% RSLogix 500 project PROGRAM 4.RSS, saved by version 8.30.00.16 %
PROJECT "UNTITLED"    % processor: Bul.1763 MicroLogix 1100 Series B %

PROGRAM FILES
  LAD 2 "MAIN"  8 rungs
  LAD 3 "IO"  7 rungs
  LAD 4 "CONTROLS"  7 rungs
  LAD 5 "CYCL_CTRL"  5 rungs
  LAD 6 "SERVO_CTRL"  4 rungs
  LAD 7 "VALVE_CTRL"  7 rungs
  LAD 8 "POS_CTRL"  6 rungs
  LAD 9 "TIMERS"  4 rungs

DATA FILES
  O0 OUTPUT  4 elements
  I1 INPUT  6 elements
  S2 STATUS  66 elements
  B3 BINARY  3 elements
  T4 TIMER  4 elements
  C5 COUNTER  1 elements
  R6 CONTROL  1 elements
  N7 INTEGER  1 elements
  F8 FLOAT  1 elements

LADDER 2 "MAIN"
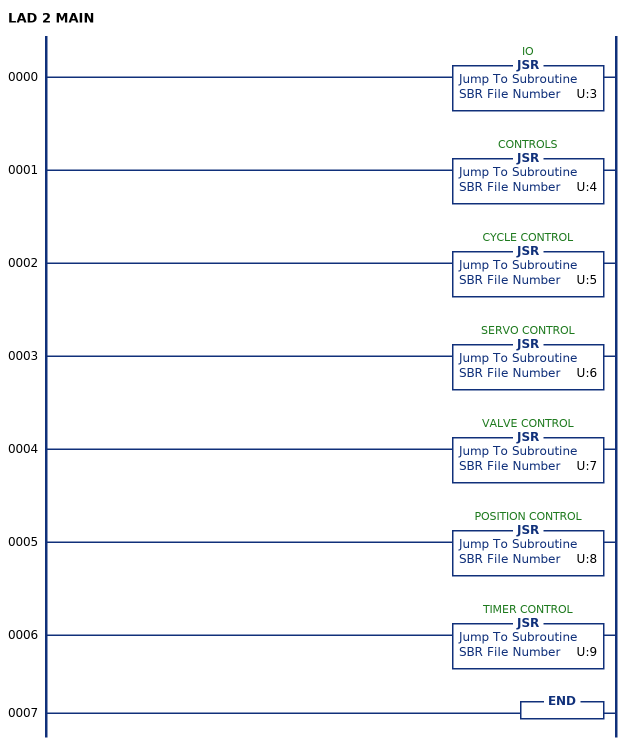
% Rung: 0 %
SOR JSR U:3 EOR
%   U:3  "IO" %
% Rung: 1 %
SOR JSR U:4 EOR
%   U:4  "CONTROLS" %
% Rung: 2 %
SOR JSR U:5 EOR
%   U:5  "CYCLE CONTROL" %
% Rung: 3 %
SOR JSR U:6 EOR
%   U:6  "SERVO CONTROL" %
% Rung: 4 %
SOR JSR U:7 EOR
%   U:7  "VALVE CONTROL" %
% Rung: 5 %
SOR JSR U:8 EOR
%   U:8  "POSITION CONTROL" %
% Rung: 6 %
SOR JSR U:9 EOR
%   U:9  "TIMER CONTROL" %
% Rung: 7 %
SOR END EOR

LADDER 3 "IO"
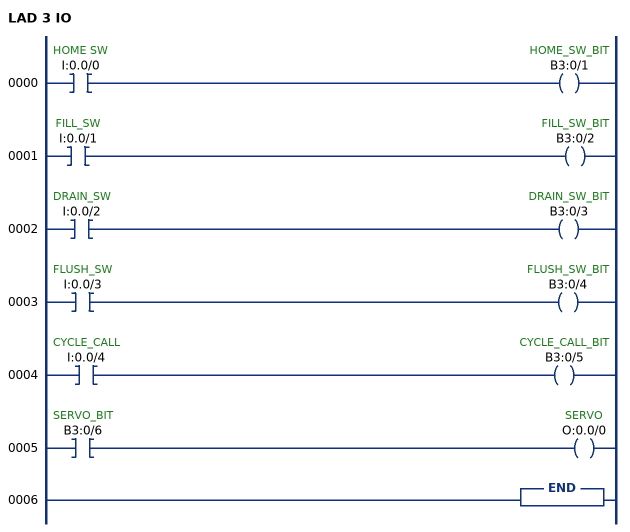
% Rung: 0 %
SOR XIC I:0.0/0 OTE B3:0/1 EOR
%   I:0.0/0  "HOME SW" %
%   B3:0/1  HOME_SW_BIT %
% Rung: 1 %
SOR XIC I:0.0/1 OTE B3:0/2 EOR
%   I:0.0/1  "FILL_SW" %
%   B3:0/2  FILL_SW_BIT %
% Rung: 2 %
SOR XIC I:0.0/2 OTE B3:0/3 EOR
%   I:0.0/2  "DRAIN_SW" %
%   B3:0/3  DRAIN_SW_BIT %
% Rung: 3 %
SOR XIC I:0.0/3 OTE B3:0/4 EOR
%   I:0.0/3  "FLUSH_SW" %
%   B3:0/4  FLUSH_SW_BIT %
% Rung: 4 %
SOR XIC I:0.0/4 OTE B3:0/5 EOR
%   I:0.0/4  "CYCLE_CALL" %
%   B3:0/5  CYCLE_CALL_BIT %
% Rung: 5 %
SOR XIC B3:0/6 OTE O:0.0/0 EOR
%   B3:0/6  SERVO_BIT %
%   O:0.0/0  "SERVO" %
% Rung: 6 %
SOR END EOR

LADDER 4 "CONTROLS"
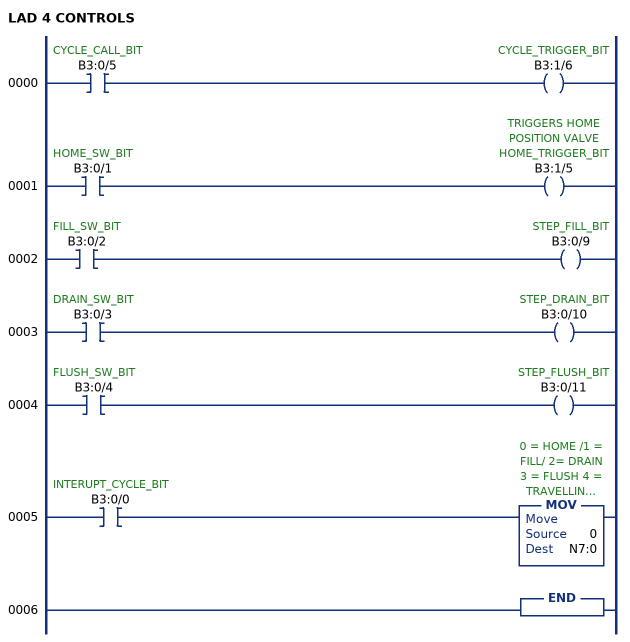
% Rung: 0 %
SOR XIC B3:0/5 OTE B3:1/6 EOR
%   B3:0/5  CYCLE_CALL_BIT %
%   B3:1/6  CYCLE_TRIGGER_BIT %
% Rung: 1 %
SOR XIC B3:0/1 OTE B3:1/5 EOR
%   B3:0/1  HOME_SW_BIT %
%   B3:1/5  HOME_TRIGGER_BIT  "TRIGGERS HOME POSITION VALVE" %
% Rung: 2 %
SOR XIC B3:0/2 OTE B3:0/9 EOR
%   B3:0/2  FILL_SW_BIT %
%   B3:0/9  STEP_FILL_BIT %
% Rung: 3 %
SOR XIC B3:0/3 OTE B3:0/10 EOR
%   B3:0/3  DRAIN_SW_BIT %
%   B3:0/10  STEP_DRAIN_BIT %
% Rung: 4 %
SOR XIC B3:0/4 OTE B3:0/11 EOR
%   B3:0/4  FLUSH_SW_BIT %
%   B3:0/11  STEP_FLUSH_BIT %
% Rung: 5 %
SOR XIC B3:0/0 MOV 0 N7:0 EOR
%   B3:0/0  INTERUPT_CYCLE_BIT %
%   N7:0  VALVE_POSITION  "0 = HOME /1 = FILL/ 2= DRAIN 3 = FLUSH 4 = TRAVELLING" %
% Rung: 6 %
SOR END EOR

LADDER 5 "CYCL_CTRL"
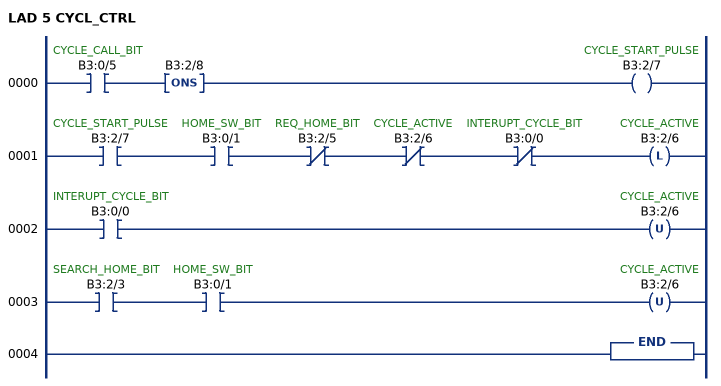
% Rung: 0 %
SOR XIC B3:0/5 ONS B3:2/8 OTE B3:2/7 EOR
%   B3:0/5  CYCLE_CALL_BIT %
%   B3:2/7  CYCLE_START_PULSE %
% Rung: 1 %
SOR XIC B3:2/7 XIC B3:0/1 XIO B3:2/5 XIO B3:2/6 XIO B3:0/0 OTL B3:2/6 EOR
%   B3:2/7  CYCLE_START_PULSE %
%   B3:0/1  HOME_SW_BIT %
%   B3:2/5  REQ_HOME_BIT %
%   B3:2/6  CYCLE_ACTIVE %
%   B3:0/0  INTERUPT_CYCLE_BIT %
% Rung: 2 %
SOR XIC B3:0/0 OTU B3:2/6 EOR
%   B3:0/0  INTERUPT_CYCLE_BIT %
%   B3:2/6  CYCLE_ACTIVE %
% Rung: 3 %
SOR XIC B3:2/3 XIC B3:0/1 OTU B3:2/6 EOR
%   B3:2/3  SEARCH_HOME_BIT %
%   B3:0/1  HOME_SW_BIT %
%   B3:2/6  CYCLE_ACTIVE %
% Rung: 4 %
SOR END EOR

LADDER 6 "SERVO_CTRL"
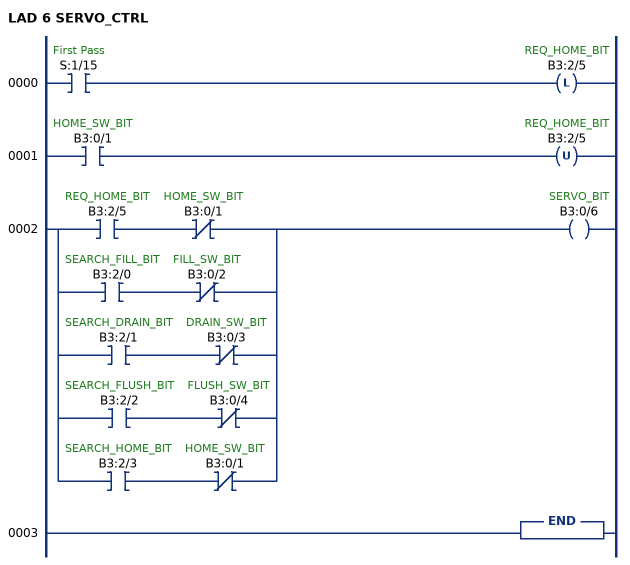
% Rung: 0 %
SOR XIC S:1/15 OTL B3:2/5 EOR
%   S:1/15  "First Pass" %
%   B3:2/5  REQ_HOME_BIT %
% Rung: 1 %
SOR XIC B3:0/1 OTU B3:2/5 EOR
%   B3:0/1  HOME_SW_BIT %
%   B3:2/5  REQ_HOME_BIT %
% Rung: 2 %
SOR BST XIC B3:2/5 XIO B3:0/1 NXB XIC B3:2/0 XIO B3:0/2 NXB XIC B3:2/1 XIO B3:0/3 NXB XIC B3:2/2 XIO B3:0/4 NXB XIC B3:2/3 XIO B3:0/1 BND OTE B3:0/6 EOR
%   B3:2/5  REQ_HOME_BIT %
%   B3:0/1  HOME_SW_BIT %
%   B3:2/0  SEARCH_FILL_BIT %
%   B3:0/2  FILL_SW_BIT %
%   B3:2/1  SEARCH_DRAIN_BIT %
%   B3:0/3  DRAIN_SW_BIT %
%   B3:2/2  SEARCH_FLUSH_BIT %
%   B3:0/4  FLUSH_SW_BIT %
%   B3:2/3  SEARCH_HOME_BIT %
%   B3:0/6  SERVO_BIT %
% Rung: 3 %
SOR END EOR

LADDER 7 "VALVE_CTRL"
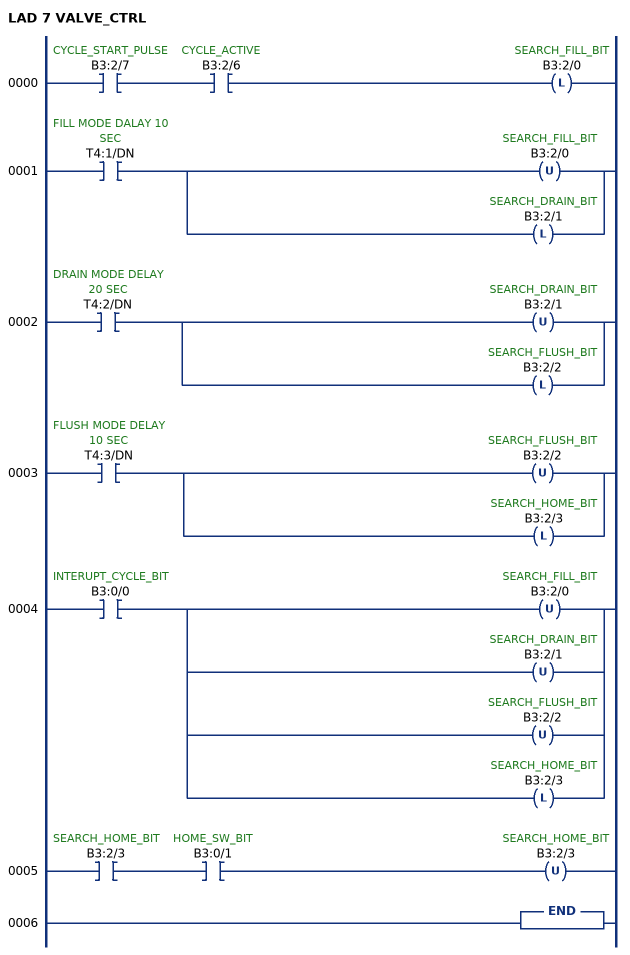
% Rung: 0 %
SOR XIC B3:2/7 XIC B3:2/6 OTL B3:2/0 EOR
%   B3:2/7  CYCLE_START_PULSE %
%   B3:2/6  CYCLE_ACTIVE %
%   B3:2/0  SEARCH_FILL_BIT %
% Rung: 1 %
SOR XIC T4:1/DN BST OTU B3:2/0 NXB OTL B3:2/1 BND EOR
%   T4:1  "FILL MODE DALAY 10 SEC" %
%   B3:2/0  SEARCH_FILL_BIT %
%   B3:2/1  SEARCH_DRAIN_BIT %
% Rung: 2 %
SOR XIC T4:2/DN BST OTU B3:2/1 NXB OTL B3:2/2 BND EOR
%   T4:2  "DRAIN MODE DELAY 20 SEC" %
%   B3:2/1  SEARCH_DRAIN_BIT %
%   B3:2/2  SEARCH_FLUSH_BIT %
% Rung: 3 %
SOR XIC T4:3/DN BST OTU B3:2/2 NXB OTL B3:2/3 BND EOR
%   T4:3  "FLUSH MODE DELAY 10 SEC" %
%   B3:2/2  SEARCH_FLUSH_BIT %
%   B3:2/3  SEARCH_HOME_BIT %
% Rung: 4 %
SOR XIC B3:0/0 BST OTU B3:2/0 NXB OTU B3:2/1 NXB OTU B3:2/2 NXB OTL B3:2/3 BND EOR
%   B3:0/0  INTERUPT_CYCLE_BIT %
%   B3:2/0  SEARCH_FILL_BIT %
%   B3:2/1  SEARCH_DRAIN_BIT %
%   B3:2/2  SEARCH_FLUSH_BIT %
%   B3:2/3  SEARCH_HOME_BIT %
% Rung: 5 %
SOR XIC B3:2/3 XIC B3:0/1 OTU B3:2/3 EOR
%   B3:2/3  SEARCH_HOME_BIT %
%   B3:0/1  HOME_SW_BIT %
% Rung: 6 %
SOR END EOR

LADDER 8 "POS_CTRL"
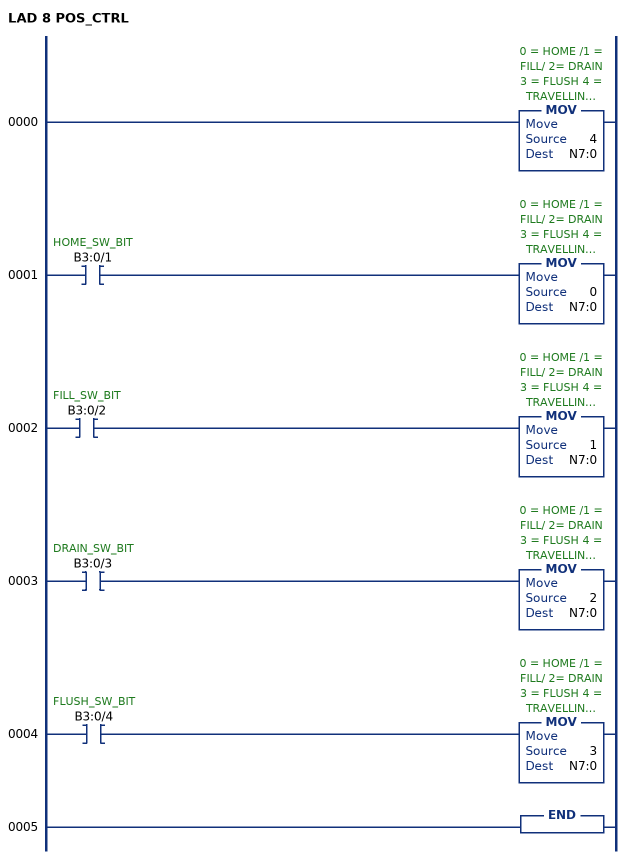
% Rung: 0 %
SOR MOV 4 N7:0 EOR
%   N7:0  VALVE_POSITION  "0 = HOME /1 = FILL/ 2= DRAIN 3 = FLUSH 4 = TRAVELLING" %
% Rung: 1 %
SOR XIC B3:0/1 MOV 0 N7:0 EOR
%   B3:0/1  HOME_SW_BIT %
%   N7:0  VALVE_POSITION  "0 = HOME /1 = FILL/ 2= DRAIN 3 = FLUSH 4 = TRAVELLING" %
% Rung: 2 %
SOR XIC B3:0/2 MOV 1 N7:0 EOR
%   B3:0/2  FILL_SW_BIT %
%   N7:0  VALVE_POSITION  "0 = HOME /1 = FILL/ 2= DRAIN 3 = FLUSH 4 = TRAVELLING" %
% Rung: 3 %
SOR XIC B3:0/3 MOV 2 N7:0 EOR
%   B3:0/3  DRAIN_SW_BIT %
%   N7:0  VALVE_POSITION  "0 = HOME /1 = FILL/ 2= DRAIN 3 = FLUSH 4 = TRAVELLING" %
% Rung: 4 %
SOR XIC B3:0/4 MOV 3 N7:0 EOR
%   B3:0/4  FLUSH_SW_BIT %
%   N7:0  VALVE_POSITION  "0 = HOME /1 = FILL/ 2= DRAIN 3 = FLUSH 4 = TRAVELLING" %
% Rung: 5 %
SOR END EOR

LADDER 9 "TIMERS"
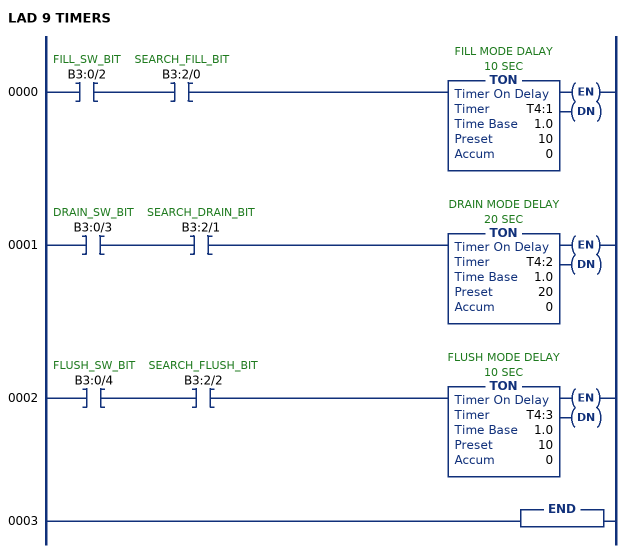
% Rung: 0 %
SOR XIC B3:0/2 XIC B3:2/0 TON T4:1 1.0 10 0 EOR
%   B3:0/2  FILL_SW_BIT %
%   B3:2/0  SEARCH_FILL_BIT %
%   T4:1  "FILL MODE DALAY 10 SEC" %
% Rung: 1 %
SOR XIC B3:0/3 XIC B3:2/1 TON T4:2 1.0 20 0 EOR
%   B3:0/3  DRAIN_SW_BIT %
%   B3:2/1  SEARCH_DRAIN_BIT %
%   T4:2  "DRAIN MODE DELAY 20 SEC" %
% Rung: 2 %
SOR XIC B3:0/4 XIC B3:2/2 TON T4:3 1.0 10 0 EOR
%   B3:0/4  FLUSH_SW_BIT %
%   B3:2/2  SEARCH_FLUSH_BIT %
%   T4:3  "FLUSH MODE DELAY 10 SEC" %
% Rung: 3 %
SOR END EOR

OTHER DOCUMENTED ADDRESSES
  B3:0/7  "HOME_SW_TRIGGER"
  B3:0/8  "FILL TRIGGER BIT"
  B3:1/0  CYCLE_ACTIVE_BIT  "OPENS CYCLE"
  B3:1/1  CYCLE_DONE_BIT  "CLOSES CYCLE"
  B3:1/2  "FILL_TRIGGER_BIT"
  B3:1/3  "DRAIN_TRIGGER_BIT"
  B3:1/4  "FLUSH_TRIGGER_BIT"
  B3:1/7  TRAVEL_BIT  "INDICATES BETWEEEN POSITION FLOW"
  C5:0  "FILL COUNTER"
  T4:0  "CYCLE CALL DELAY"
  T4:1/EN  "BETWEEN POSTIONS"

DATA TABLE (non-zero values as saved)
DATA T4
% .PRE .ACC %
% T4:1 % 10 0
% T4:2 % 20 0
% T4:3 % 10 0
